(*
SPDX-FileCopyrightText: © 2026 Oleksandr Tiutyk <trofimich@gmail.com>
SPDX-License-Identifier: MIT
License: https://opensource.org/license/mit
*)

(*!
<summary>Represents an exception raised when an invalid workflow state transition is requested or attempted.</summary>
<description>
Instances are task-scoped diagnostic objects; do not retain references across PLC task cycles.
</description>
*)

INTERFACE IInvalidWorkflowTransitionException EXTENDS TOF_Core.IGeneralException

(*!
<summary>Formats the invalid state transition diagnostic and raises this exception.</summary>
<description>
Formats bounded diagnostic text without allocating temporary builder storage. Propagation follows the Core
exception lifetime and allocation rules and does not return normally in valid cyclic-task usage.
</description>
<param name="sourceNamespaceName">Namespace of the POU raising the exception.</param>
<param name="sourceClassName">Class name of the workflow element where the transition was rejected.</param>
<param name="sourcePOUName">Method or property name where the transition was attempted.</param>
<param name="sourcePosition">Source position identifier.</param>
<param name="fromState">Current state of the workflow element.</param>
<param name="toState">Rejected target state.</param>
*)
METHOD Throw
VAR_INPUT
	sourceNamespaceName : STRING;
	sourceClassName : STRING;
	sourcePOUName : STRING;
	sourcePosition : STRING;
	fromState : WORKFLOW_ELEMENT_STATE;
	toState : WORKFLOW_ELEMENT_STATE;
END_VAR
END_METHOD

END_INTERFACE

(* stored: Version 1.1.0.1
   Itf IInvalidWorkflowTransitionException: Id {7340e873-0fee-42d6-bda3-e9bfd586f0f4}
   Method Throw: Id {6c679139-20ab-4061-b94a-4c6f3303172c} *)
